// TIA Portal V20 export
Screen "Pop-up_IF_SIGNALS_LEGEND_Popup"  327x200
  ScreenItem "Background" at 0,0 size 327x200  Type=HmiRectangle
  ScreenItem "Textfeld_15" at 10,85 size 250x20  Type=HmiTextBox
  ScreenItem "Cancel Mode" at 236,1 size 90x60  Type=HmiButton
  ScreenItem "Textfeld_1" at 10,107 size 300x20  Type=HmiTextBox
  ScreenItem "Textfeld_2" at 10,132 size 250x20  Type=HmiTextBox
  ScreenItem "Textfeld_3" at 10,154 size 310x35  Type=HmiTextBox
  ScreenItem "Textfeld_4" at 10,10 size 210x75  Type=HmiTextBox
